(* IEC 61131-3 sources: Gen-AI/release/member2-v1.1/成员2_提交包_v1.1/agent/logs/full34_fixture/E3_S03_1_42/tools/candidate_1/fixture_compile, 1 file *)

(* ---- source.st ---- *)
FUNCTION_BLOCK FB_S03
VAR_INPUT
    DoorSwitch : BOOL;
    ZoneAOccupied : BOOL;
    ZoneBOccupied : BOOL;
    ResetBtn : BOOL;
    EStop_NC : BOOL;
END_VAR
VAR_OUTPUT
    DriveA_Run : BOOL;
    DriveB_Run : BOOL;
    AlarmLamp : BOOL;
    Status : WORD;
END_VAR
(* Add a VAR block for internal state/timers before the implementation, if needed. *)
(* SKELETON ONLY: replace this RETURN with scan logic and required initial state. *)
RETURN;
END_FUNCTION_BLOCK

(* FIXTURE_COMPILE_FAIL *)
